(* PLC project probe.project, CODESYS CODESYS V3.5 SP17 Patch 3 *)
(* stored: creationDateTime 2026-10-20T03:54:26.8299914, modificationDateTime 1601-01-01T03:00:00 *)

FUNCTION_BLOCK FB_ProbePcfc
  VAR_INPUT
    rA : REAL;
    rK : REAL;
  END_VAR
  VAR_OUTPUT
    rEarly : REAL;
    rLate : REAL;
  END_VAR
  VAR  (* added by the conversion: wires and edge detectors of the diagram *)
    _MUL3_OUT : ANY;
  END_VAR

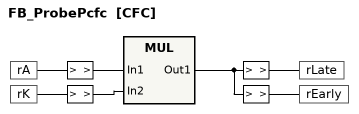
(* CFC diagram, written out as Structured Text *)
rEarly := _MUL3_OUT;
_MUL3_OUT := rA * rK;
rLate := _MUL3_OUT;
END_FUNCTION_BLOCK
